// Mitsubishi GX Works2 project: Test_Station_2   PLC: Q03UD

PROGRAM MAIN
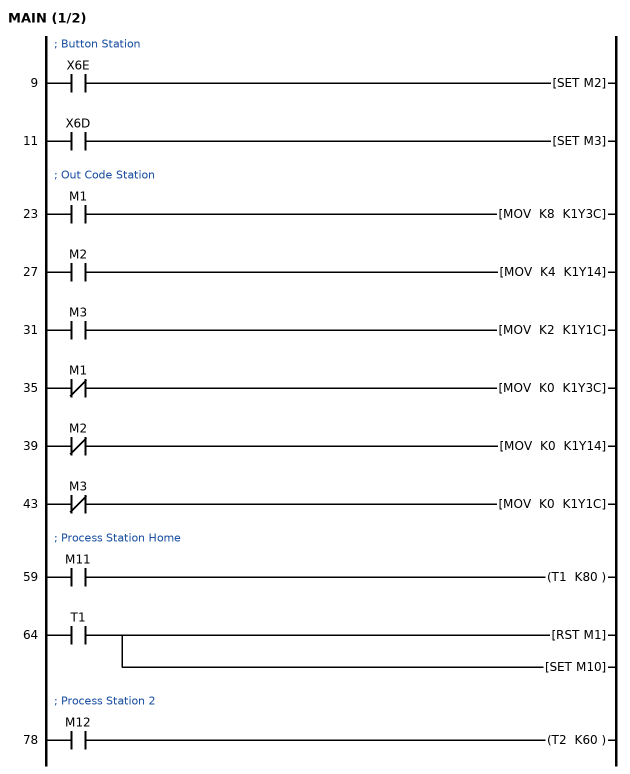
; Button Station
9     LD      X6E
      SET     M2
11    LD      X6D
      SET     M3
; Out Code Station
23    LD      M1
      MOV     K8 K1Y3C
27    LD      M2
      MOV     K4 K1Y14
31    LD      M3
      MOV     K2 K1Y1C
35    LDI     M1
      MOV     K0 K1Y3C
39    LDI     M2
      MOV     K0 K1Y14
43    LDI     M3
      MOV     K0 K1Y1C
; Process Station Home
59    LD      M11
      OUT     T1 K80
64    LD      T1
      RST     M1
      SET     M10
; Process Station 2
78    LD      M12
      OUT     T2 K60
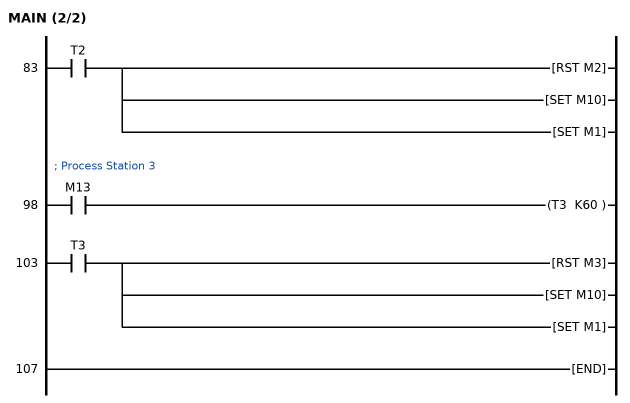
83    LD      T2
      RST     M2
      SET     M10
      SET     M1
; Process Station 3
98    LD      M13
      OUT     T3 K60
103   LD      T3
      RST     M3
      SET     M10
      SET     M1
107   END
END_PROGRAM
